(* IEC 61131-3 sources: plc-vscode/tests/st/all/trust-platform/crates/trust-runtime/tests/fixtures/plcopen_motion/single_axis_negative_stop_active/src, 2 files *)

(* ---- main.st ---- *)
PROGRAM Main
VAR
    Axis : AXIS_REF;
    Stop : MC_Stop;
END_VAR

Stop(Axis := Axis, Execute := TRUE, Deceleration := REAL#1.0, Jerk := REAL#1.0);
IF Stop.Active THEN
END_IF;
END_PROGRAM

(* ---- tests.st ---- *)
TEST_PROGRAM plcopen_motion_single_axis_negative_stop_active
VAR
    Axis : AXIS_REF;
    Stop : MC_Stop;
END_VAR

Stop(Axis := Axis, Execute := TRUE, Deceleration := REAL#1.0, Jerk := REAL#1.0);
ASSERT_FALSE(Stop.Active);
END_TEST_PROGRAM
